{attribute 'qualified_only'}
VAR_GLOBAL
    start : BOOL;
    stop : BOOL;
    guardClosed : BOOL := TRUE;
    productSensor : BOOL;
    resetCount : BOOL;
    motorRunning : BOOL;
    productCount : UDINT;
    alarm : STRING(80);
END_VAR

(* stored: Version 1.1.0.1, ProductVersion 3.1 *)
